// TIA Portal V17 export
FUNCTION_BLOCK "ValveActuator"   // FB, LAD
// Opens the pneumatic valve actuator when the open command is on and the closed feedback has dropped.
   VAR_INPUT
      OpenCommand : Bool;   // Open command
      ClosedFeedback : Bool;   // Closed feedback
   END_VAR
   VAR_OUTPUT
      Actuator : Bool;   // Pneumatic valve actuator
   END_VAR
BEGIN

REGION Network 1: Open the valve actuator
   // Fault: the valve did not leave the closed position.
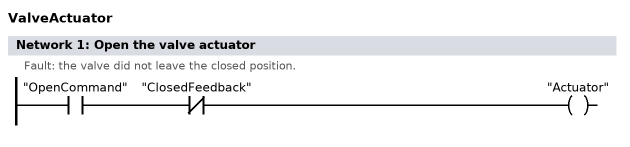
   RUNG wire#powerrail
      Contact( "OpenCommand" )
      I_Contact( "ClosedFeedback" )
      Coil( "Actuator" )
   END_RUNG
   // the same network as SCL:
   "Actuator" := "OpenCommand" AND NOT "ClosedFeedback";
END_REGION
END_FUNCTION_BLOCK
